{attribute 'qualified_only'}
VAR_GLOBAL
    bStart AT %I* : BOOL;
END_VAR

(* stored: Version 1.1.0.1
   GVL GVL_IO: Id {00000000-0000-0000-0000-000000000001} *)
